FUNCTION_BLOCK FB_ExampleStation EXTENDS FB_Module
(*
	Example station with two 2-state actuators and a trigger/tell transaction.
	Home position = OPEN, Work position = CLOSED.
	
	Starting (homing)	: open both actuators, Started once both are open
	Started (running)	: one job per cycle:
						  ask the software for a job (attention), validate and ack the request,
						  close both, hold for request.closeDwell, open both, report (tell), dwell
	Stopping			: abort any open transaction, open both actuators (safe position)
	Stopped				: actuators follow operator commands (manual mode)
	
	The actuators are configured with no feedback so the example runs without hardware.
	Clear homeNoFdbk/workNoFdbk and link homeFdbk/workFdbk/outHome/outWork to use real I/O.
*)
VAR_INPUT
	{attribute 'OPC.UA.DA' := '1'}
	{attribute 'OPC.UA.DA.StructuredType' := '1'}
	cfg					: ST_ExampleStationConfiguration; //configuration
	
	(* Devices
	----------------------------------------------------------------------------------------------------*)
	{attribute 'OPC.UA.DA' := '1'}
	actuatorA			: FB_Actuator2State := (cfg := (actuatorId := 'Actuator A', homeNoFdbk := TRUE, workNoFdbk := TRUE));
	{attribute 'OPC.UA.DA' := '1'}
	actuatorB			: FB_Actuator2State := (cfg := (actuatorId := 'Actuator B', homeNoFdbk := TRUE, workNoFdbk := TRUE));
	
	(* Communication
	----------------------------------------------------------------------------------------------------*)
	{attribute 'OPC.UA.DA' := '1'}
	transaction			: FB_ExampleTransaction := (cfg := (commTimeout := T#10S)); //job request/response with the software
END_VAR
VAR_OUTPUT
	{attribute 'OPC.UA.DA' := '1'}
	{attribute 'OPC.UA.DA.Access' := '1'}
	{attribute 'OPC.UA.DA.StructuredType' := '1'}
	stsStation			: ST_ExampleStationStatus; //station specific status (module status is in sts)
END_VAR
VAR
	//Timers
	dwellTimer			: TON; //dwell between cycles
	holdTimer			: TON; //holds the actuators closed for job.closeDwell
	cycleTimer			: TON := (PT := T#1D); //measures one close/hold/open cycle
END_VAR

SUPER^();

Devices();
Permissives();
StatusOut();

METHOD PROTECTED CloseAll //command all actuators to work (closed)
IF NOT actuatorA.sts.atWork AND NOT actuatorA.sts.goingToWork THEN
	actuatorA.ToWork();
END_IF
IF NOT actuatorB.sts.atWork AND NOT actuatorB.sts.goingToWork THEN
	actuatorB.ToWork();
END_IF
END_METHOD

METHOD PROTECTED Devices //call child devices
//Devices follow this module's mode through childCtrl
actuatorA(parentCtrl := childCtrl);
actuatorB(parentCtrl := childCtrl);
transaction();

//Report child faults to the module
inpChildFaulted := actuatorA.fault.active OR actuatorB.fault.active;
END_METHOD

METHOD PROTECTED OpenAll //command all actuators to home (open)
IF NOT actuatorA.sts.atHome AND NOT actuatorA.sts.goingToHome THEN
	actuatorA.ToHome();
END_IF
IF NOT actuatorB.sts.atHome AND NOT actuatorB.sts.goingToHome THEN
	actuatorB.ToHome();
END_IF
END_METHOD

METHOD PROTECTED Permissives //set module permissives and interlocks
//Homing is complete when all actuators are open
PermStartComplete.cfg.condText[0] := 'Actuator A open';
PermStartComplete.cfg.condText[1] := 'Actuator B open';
PermStartComplete.perm.0 := actuatorA.sts.atHome;
PermStartComplete.perm.1 := actuatorB.sts.atHome;

//Stopping is complete when all actuators are open, or faulted so they cannot move
PermStopComplete.cfg.condText[0] := 'Actuator A open or faulted';
PermStopComplete.cfg.condText[1] := 'Actuator B open or faulted';
PermStopComplete.perm.0 := actuatorA.sts.atHome OR actuatorA.fault.active;
PermStopComplete.perm.1 := actuatorB.sts.atHome OR actuatorB.fault.active;

//A faulted actuator stops the station
IntlkAuto.cfg.condText[0] := 'Actuator A not faulted';
IntlkAuto.cfg.condText[1] := 'Actuator B not faulted';
IntlkAuto.perm.0 := NOT actuatorA.fault.active;
IntlkAuto.perm.1 := NOT actuatorB.fault.active;
END_METHOD

METHOD PUBLIC Reset : BOOL
actuatorA.Reset();
actuatorB.Reset();
transaction.Reset();
Reset := TRUE;
END_METHOD

METHOD PROTECTED Started : BOOL
//Running sequence: one trigger/tell transaction per close/open cycle
CASE stsStation.runStep OF
	
	E_ExampleStationRunStep.Idle:
		stsStation.runStep := E_ExampleStationRunStep.RequestJob;
		
	E_ExampleStationRunStep.RequestJob:
		IF transaction.sts.Idle THEN
			transaction.Start(); //raises attention
			stsStation.runStep := E_ExampleStationRunStep.WaitJob;
		END_IF
		
	E_ExampleStationRunStep.WaitJob:
		IF transaction.sts.Request_Start THEN
			IF ValidateJob(transaction.request) THEN
				stsStation.job := transaction.request;
				transaction.SetRequestACK();
				stsStation.runStep := E_ExampleStationRunStep.WaitWorking;
			ELSE
				transaction.Abort();
				stsStation.jobsRejected := stsStation.jobsRejected + 1;
				stsStation.runStep := E_ExampleStationRunStep.Dwell;
			END_IF
		END_IF
		
	E_ExampleStationRunStep.WaitWorking:
		IF transaction.sts.Working THEN
			stsStation.runStep := E_ExampleStationRunStep.Close;
		END_IF
		
	E_ExampleStationRunStep.Close:
		CloseAll();
		IF stsStation.allClosed THEN
			stsStation.runStep := E_ExampleStationRunStep.HoldClosed;
		END_IF
		
	E_ExampleStationRunStep.HoldClosed:
		IF holdTimer.Q THEN
			stsStation.runStep := E_ExampleStationRunStep.Open;
		END_IF
		
	E_ExampleStationRunStep.Open:
		OpenAll();
		IF stsStation.allOpen THEN
			stsStation.lastCycleTime := cycleTimer.ET;
			stsStation.runStep := E_ExampleStationRunStep.Report;
		END_IF
		
	E_ExampleStationRunStep.Report:
		transaction.response.cycleId 	:= stsStation.job.cycleId;
		transaction.response.cycleTime 	:= stsStation.lastCycleTime;
		transaction.response.ok 		:= NOT (actuatorA.fault.active OR actuatorB.fault.active);
		transaction.FinishWork(); //raises tell
		stsStation.cycleCount := stsStation.cycleCount + 1;
		stsStation.runStep := E_ExampleStationRunStep.WaitReportAck;
		
	E_ExampleStationRunStep.WaitReportAck:
		IF transaction.sts.Idle THEN
			stsStation.runStep := E_ExampleStationRunStep.Dwell;
		END_IF
		
	E_ExampleStationRunStep.Dwell:
		IF dwellTimer.Q THEN
			stsStation.runStep := E_ExampleStationRunStep.RequestJob;
		END_IF
		
END_CASE
END_METHOD

METHOD PROTECTED Starting : BOOL
//Homing: open all actuators, no transaction open
OpenAll();
AbortTransaction();
stsStation.runStep := E_ExampleStationRunStep.Idle;
END_METHOD

METHOD PROTECTED StatusOut //Set output status information
stsStation.allOpen 	:= actuatorA.sts.atHome AND actuatorB.sts.atHome;
stsStation.allClosed 	:= actuatorA.sts.atWork AND actuatorB.sts.atWork;

stsStation.commError 	:= transaction.sts.errTimeout;

//Monitoring timers
dwellTimer(IN := stsStation.runStep = E_ExampleStationRunStep.Dwell, PT := cfg.cycleDwell);
holdTimer(IN := stsStation.runStep = E_ExampleStationRunStep.HoldClosed, PT := stsStation.job.closeDwell);
cycleTimer(IN := stsStation.runStep = E_ExampleStationRunStep.Close
			OR stsStation.runStep = E_ExampleStationRunStep.HoldClosed
			OR stsStation.runStep = E_ExampleStationRunStep.Open);
END_METHOD

METHOD PROTECTED Stopping : BOOL
//Finish in the safe position: all actuators open, transaction closed
OpenAll();
AbortTransaction();
stsStation.runStep := E_ExampleStationRunStep.Idle;
END_METHOD

METHOD PROTECTED AbortTransaction //cancel an open transaction
IF transaction.sts.bBusy THEN
	transaction.Abort();
END_IF
END_METHOD

METHOD PROTECTED ValidateJob : BOOL //TRUE if the request can be worked on, sets lastRejectText otherwise
VAR_INPUT
	job			: ST_ExampleRequest;
END_VAR
IF job.closeDwell <= T#0S THEN
	stsStation.lastRejectText := 'closeDwell must be greater than 0';
ELSIF job.closeDwell > cfg.maxCloseDwell THEN
	stsStation.lastRejectText := 'closeDwell is longer than cfg.maxCloseDwell';
ELSE
	ValidateJob := TRUE;
	RETURN;
END_IF
ValidateJob := FALSE;
END_METHOD

END_FUNCTION_BLOCK

(* stored: Version 1.1.0.1, ProductVersion 3.1.4024.12
   POU FB_ExampleStation: Id {ec9942f8-1fba-4f7b-ba35-139c4983ee10}, SpecialFunc None
   Folder Protected: Id {e23fc091-61a6-4328-b2d5-222d594dc1f8}
   Folder Logic: Id {eae64112-d142-48a0-b521-dc602e636cee}
   Folder States: Id {78beda1c-b282-44b8-97c0-52fabcb170bf}
   Folder Public: Id {a38f987d-ca93-474e-ab80-c214117163e7}
   Folder Control: Id {945794ed-2e4e-4654-93eb-8e546ac0d6eb}
   Method CloseAll: Id {8e52d248-87df-4c42-99f6-9d9c54f47983}
   Method Devices: Id {f44671b1-c0e4-43be-93bd-be3677fe4079}
   Method OpenAll: Id {1e08200a-bb87-4855-85ad-e602e4fc47d6}
   Method Permissives: Id {d88cb704-047f-4a29-9dd2-a0bdee56da70}
   Method Reset: Id {23c61360-e642-4960-8caa-c42cb99c1793}
   Method Started: Id {766cf290-1a71-461d-81fe-613336b7212d}
   Method Starting: Id {3fe50c0b-caad-4b2b-8963-ca5f99eef799}
   Method StatusOut: Id {9145cda4-cd6c-47f3-90f1-a708e1e13d88}
   Method Stopping: Id {51f6e602-e616-41ff-b9af-086d08317e64}
   Method AbortTransaction: Id {0f8ac1c9-2c94-41b9-873e-b37a0981dad2}
   Method ValidateJob: Id {8c3e32c7-7e51-442c-ad45-d75788e1cd57} *)
